(* PLC project station_cds.project, CODESYS CODESYS V3.5 SP22 Patch 1 *)
(* stored: creationDateTime 2026-11-25T17:27:32.3706002, modificationDateTime 2026-11-25T17:27:31.3827148 *)

FUNCTION_BLOCK FB_TestPlant
  VAR_INPUT
    Reset : BOOL;  (* a new part is in the fixture *)
    CycleTime : REAL := 0.002;  (* s *)
    QVel : REAL;  (* mm/s *)
    QDriveEnable : BOOL;
    QClamp : BOOL;
    PartPresent : BOOL;
    Curve : INT;  (* recorded curve the part follows *)
    Seat : REAL := 5.0;  (* mm, axis position at which the hook meets the grip *)
  END_VAR
  VAR_OUTPUT
    Pos : REAL;  (* mm *)
    Force : REAL;  (* N *)
    ClampClosed : BOOL;
    ClampOpen : BOOL;
    Moved : BOOL;  (* the axis has moved or the clamp has closed since the last Reset *)
  END_VAR
  VAR
    sPos : REAL;
    sClamp : REAL;
    sReturn : BOOL;
    sK : INT;
    sMoved : BOOL;
  END_VAR
  VAR_TEMP
    tI : INT;
    tA : INT;
    tN : INT;
    tX : REAL;
    tF : REAL;
    tX0 : REAL;
    tX1 : REAL;
    tF0 : REAL;
    tF1 : REAL;
  END_VAR

                {region "Part"}
        IF Reset THEN
            sReturn := FALSE;
            sK := 0;
            sMoved := FALSE;
        END_IF;
    {endregion}

    {region "AxisAndClamp"}
        IF QDriveEnable THEN
            sPos := sPos + QVel * CycleTime;
            IF QVel <> 0.0 THEN
                sMoved := TRUE;
            END_IF;
        END_IF;
        IF sPos < 0.0 THEN
            sPos := 0.0;
        END_IF;
        IF QClamp THEN
            sClamp := sClamp + CycleTime;
            sMoved := TRUE;
        ELSE
            sClamp := sClamp - CycleTime;
        END_IF;
        sClamp := LIMIT(0.0, sClamp, 0.25);
    {endregion}

    {region "Handle"}
        tX := sPos - Seat;
        tF := 0.0;
        tA := GVL_TestData.CurveStart[Curve];
        tN := GVL_TestData.CurveNPull[Curve];
        IF QVel < 0.0 AND NOT sReturn THEN
            sReturn := TRUE;
            sK := 0;
        END_IF;
        IF PartPresent AND tX >= 0.0 AND tN >= 2 THEN
            IF sReturn THEN
                tA := tA + tN;   // the return samples follow the pull samples; their travel falls
            END_IF;
            // move on to the pair of samples around the travel (the axis moves less than 8 samples per call)
            FOR tI := 1 TO 8 DO
                IF sK < tN - 2 THEN
                    IF NOT sReturn AND GVL_TestData.X[tA + sK + 1] < tX THEN
                        sK := sK + 1;
                    ELSIF sReturn AND GVL_TestData.X[tA + sK + 1] > tX THEN
                        sK := sK + 1;
                    END_IF;
                END_IF;
            END_FOR;
            tX0 := GVL_TestData.X[tA + sK];
            tX1 := GVL_TestData.X[tA + sK + 1];
            tF0 := GVL_TestData.F[tA + sK];
            tF1 := GVL_TestData.F[tA + sK + 1];
            IF NOT sReturn THEN
                IF tX >= tX1 THEN
                    tF := tF1 + (tX - tX1) * 25.0;
                ELSIF tX <= tX0 OR tX1 - tX0 < 0.000001 THEN
                    tF := tF0;
                ELSE
                    tF := tF0 + (tF1 - tF0) * (tX - tX0) / (tX1 - tX0);
                END_IF;
            ELSE
                IF tX >= tX0 THEN
                    tF := tF0 + (tX - tX0) * 25.0;
                ELSIF tX <= tX1 OR tX0 - tX1 < 0.000001 THEN
                    tF := tF1;
                ELSE
                    tF := tF1 + (tF0 - tF1) * (tX - tX1) / (tX0 - tX1);
                END_IF;
            END_IF;
        END_IF;
    {endregion}

    {region "Outputs"}
        Pos := sPos;
        Force := tF;
        ClampClosed := sClamp >= 0.25;
        ClampOpen := sClamp <= 0.0;
        Moved := sMoved;
    {endregion}

          
END_FUNCTION_BLOCK
